(* IEC 61131-3 sources: JingjiangArm/moonboxpro_arm_8.4/Application/Application/任务列表/CommTask/轴号站号处理, 8 files *)

(* ---- KS_CheckArcIdValid.st ---- *)
(*@CES
Name=KS_CheckArcIdValid
Type=FunctionBlock
TypeGuid=6f9dac99-8de1-4efc-8465-68ac443b7d08
Guid=246184da-21c6-48ff-adc4-5d24f4660108
HasDeclaration=True
HasImplementation=True
*)
{DECLARATION}
FUNCTION KS_CheckArcIdValid : BOOL
VAR_INPUT
	i_iAxisId:INT;(*轴id*)
	i_iArcId:INT;(*套色id@修改后的*)
	i_pabyColorIdCurrent: POINTER TO ARRAY [1..MAX_UNIT_NUM] OF BYTE;(*色组色序*)
END_VAR
VAR
	iN: INT;
	xValid:BOOL:=TRUE;(*默认是有效的*)
END_VAR

{IMPLEMENTATION}
IF i_pabyColorIdCurrent<>0 THEN
	IF i_iAxisId>1 AND i_iArcId>1 THEN
		FOR iN:=1 TO i_iAxisId-1 BY 1 DO(*检查修改的轴前面的轴套色id*)
			IF i_pabyColorIdCurrent^[iN]>1 THEN(**)
				IF i_iArcId>i_pabyColorIdCurrent^[iN] THEN(*新修改的比上面轴的大就行*);
				ELSE(*小于等于任何一个都认为是无效的*)
					xValid:=FALSE;
					EXIT;
				END_IF
			END_IF
		END_FOR
	END_IF
END_IF

KS_CheckArcIdValid:=xValid;

(* ---- KS_GetArcIdList.st ---- *)
(*@CES
Name=KS_GetArcIdList
Type=FunctionBlock
TypeGuid=6f9dac99-8de1-4efc-8465-68ac443b7d08
Guid=d22e29e8-5d32-4a53-8a83-de107a05006d
HasDeclaration=True
HasImplementation=True
*)
{DECLARATION}
FUNCTION KS_GetArcIdList : BOOL
VAR_INPUT
	i_xEn:BOOL;(*更新列表使能标志*)
	i_iGrpAxisNum_Pu: INT; (*系的轴数量*)
	i_aiGrpAxisList: ARRAY [1..MAX_UNIT_NUM] OF INT; (*系的轴列表|已经按照升序排列了*)
	i_paxArcEnSts_Bak:POINTER TO ARRAY [1..MAX_UNIT_NUM] OF BOOL;(*套色使能备份值|用于检查是否套色使能切换*)
	i_pabyArcId_Bak:POINTER TO ARRAY [1..MAX_UNIT_NUM] OF BYTE;(*备份套色id*)
	(*系套色轴个数@可以输入0*)
	i_piGrpArcAxisNum_Pu:POINTER TO INT;
	i_axLinkage: ARRAY [1..MAX_UNIT_NUM] OF BOOL;
	i_axThisUnitEna: ARRAY [1..MAX_UNIT_NUM] OF BOOL;
	i_axSwitchOn_CoatingPrn: ARRAY [1..MAX_UNIT_NUM] OF BOOL;
	i_pabyColorIdCurrent: POINTER TO ARRAY [1..MAX_UNIT_NUM] OF BYTE;(*色组色序*)

END_VAR
VAR
	iN:INT;
	iUnitId:INT;
	xArcEnSts:BOOL;(*套色使能值|用于检查是否套色使能切换*)
	axArcEnSts_Bak:ARRAY [1..MAX_UNIT_NUM] OF BOOL;(*套色使能备份值|用于检查是否套色使能切换*)
	abyArcId_Bak:ARRAY [1..MAX_UNIT_NUM] OF BYTE;(*备份套色id*)
	(*系套色个数*)
	iGrpArcAxisNum_Pu:INT;
	xNeedUpdate: BOOL;
	byAxisIdArcValid: BYTE;(*最后一个未更新套色id|有效的轴id*)
	iAxisIdSa_Update: INT;(*更新的起始id@后面轴的套色id都更新*)
	xArcIdLocked:BOOL;(*套色id被锁定了|在更新的时候不修改这个值*)
	xRtn: BOOL;
	xUpdateArcId_BakValue: BOOL;(*更新套色id的备份值*)
	iIndex: INT;
END_VAR

{IMPLEMENTATION}
IF i_paxArcEnSts_Bak<>0 AND
	i_pabyArcId_Bak<>0 AND
	i_pabyColorIdCurrent<>0 THEN

	IF i_xEn THEN
		axArcEnSts_Bak:=i_paxArcEnSts_Bak^;(*获取之前的备份值*)
		abyArcId_Bak:=i_pabyArcId_Bak^;(*备份套色id*)

		FOR iN:=1 TO i_iGrpAxisNum_Pu BY 1 DO
			iUnitId:=i_aiGrpAxisList[iN];

			xArcEnSts:=i_axThisUnitEna[iUnitId] AND(*使能了*)
				i_axLinkage[iUnitId] AND(*联动了*)
				(NOT i_axSwitchOn_CoatingPrn[iUnitId]);(*不是涂布色组*)

			IF xArcEnSts<>axArcEnSts_Bak[iUnitId] THEN(*有轴的状态发生变化了*)
				IF NOT xNeedUpdate THEN(*记录需要更新的开始轴id*)
					iAxisIdSa_Update:=iUnitId;
				END_IF
				xNeedUpdate:=TRUE;
			END_IF

			(*记录最后一个不更新套色id的轴*)
			IF NOT xNeedUpdate THEN(*还没找到需要变化的轴id*)
				IF i_pabyColorIdCurrent^[iUnitId]<>0 THEN
					byAxisIdArcValid:= i_pabyColorIdCurrent^[iUnitId];
				END_IF
			END_IF
			axArcEnSts_Bak[iUnitId]:=xArcEnSts;
		END_FOR

		IF NOT xNeedUpdate THEN(*手动更新列表@注意调用顺序*)
			FOR iN:=1 TO i_iGrpAxisNum_Pu BY 1 DO
				iUnitId:=i_aiGrpAxisList[iN];
				xArcEnSts:=axArcEnSts_Bak[iUnitId];
				IF NOT xArcEnSts THEN(*套色不使能的时候 手动也不能输入*)
					i_pabyColorIdCurrent^[iUnitId]:=0;(*强制写0*)
				ELSE
					IF i_pabyColorIdCurrent^[iUnitId]=0 THEN(*输入了0则强制写成备份值*)
						i_pabyColorIdCurrent^[iUnitId]:=abyArcId_Bak[iUnitId];
						EXIT;(*手动修改了*)
					ELSE
						IF abyArcId_Bak[iUnitId]<>i_pabyColorIdCurrent^[iUnitId] THEN(*id被修改了*)
							xRtn:=KS_CheckArcIdValid(iUnitId,i_pabyColorIdCurrent^[iUnitId],i_pabyColorIdCurrent);
							IF xRtn THEN(*id合法@手动修改成功了|后面的列表需要同步更新*)
								xNeedUpdate:=TRUE;(*由下面逻辑生成*)
								iAxisIdSa_Update:=iUnitId;
								byAxisIdArcValid:=i_pabyColorIdCurrent^[iUnitId]-1;(*更新的时候会+1*)
							ELSE(*不合法@保持之前的*)
								i_pabyColorIdCurrent^[iUnitId]:=abyArcId_Bak[iUnitId];
							END_IF
							(*pstStAxisParam^.byColorIdCurrent 界面修改的,不在同一个任务中,防止不能抓住改变的状态
							置标志只有进入过这里才更新备份值*)
							xUpdateArcId_BakValue:=TRUE;

							EXIT;(*手动修改了*)
						END_IF
					END_IF
				END_IF
			END_FOR
		END_IF

		(*上面执行完成后axArcEnSts_Bak 中存储的每个色组是否套色的状态*)
		IF xNeedUpdate THEN(*自动更新列表了*)
			(*套色轴个数初始化*)
			IF byAxisIdArcValid<>0 THEN
				iGrpArcAxisNum_Pu:=BYTE_TO_INT(byAxisIdArcValid);
			ELSE
				iGrpArcAxisNum_Pu:=0;
			END_IF

			(*找到起始轴的索引值*)
			FOR iN:=1 TO i_iGrpAxisNum_Pu BY 1 DO
				iUnitId:=i_aiGrpAxisList[iN];
				IF iAxisIdSa_Update = iUnitId THEN
					iIndex:=iN;
					EXIT;
				END_IF
			END_FOR

			FOR iN:=iIndex TO i_iGrpAxisNum_Pu BY 1 DO(*从变化的轴这里开始，更新后面的套色id*)
				iUnitId:=i_aiGrpAxisList[iN];
				xArcEnSts:=axArcEnSts_Bak[iUnitId];

//xArcIdLocked;(*还未处理*)

				IF xArcEnSts THEN(*套色使能了*)
					iGrpArcAxisNum_Pu:=iGrpArcAxisNum_Pu+1;
					IF NOT xArcIdLocked THEN(*套色Id未被锁定*)
						i_pabyColorIdCurrent^[iUnitId]:=INT_TO_BYTE(iGrpArcAxisNum_Pu);
					ELSE(*套色Id被锁定了|当前色序id不做修改,更新套色轴个数变量*)
						IF i_pabyColorIdCurrent^[iUnitId]>iGrpArcAxisNum_Pu THEN
							iGrpArcAxisNum_Pu:=i_pabyColorIdCurrent^[iUnitId];
						ELSE
							i_pabyColorIdCurrent^[iUnitId]:=INT_TO_BYTE(iGrpArcAxisNum_Pu);
						END_IF
					END_IF
				ELSE
					i_pabyColorIdCurrent^[iUnitId]:=0;
				END_IF
			END_FOR
		ELSE(*在不更新的时候支持手动的输入*);
		END_IF

		(*更新存储的备份值@不用做专门的备份值初始化,因为刚上电的大概率肯定会更新列表*)
		FOR iN:=1 TO i_iGrpAxisNum_Pu BY 1 DO
			iUnitId:=i_aiGrpAxisList[iN];
			(*pstStAxisParam^.byColorIdCurrent 界面修改的,不在同一个任务中,防止不能抓住改变的状态
			置标志只有进入过上面逻辑更新备份值*)
			IF xUpdateArcId_BakValue OR xNeedUpdate THEN(*或者更新了列表后就更新*)
				abyArcId_Bak[iUnitId]:=i_pabyColorIdCurrent^[iUnitId];
			END_IF
		END_FOR
	ELSE;(*不使能*)
	END_IF

	i_paxArcEnSts_Bak^:=axArcEnSts_Bak;(*更新备份值|en=false 全部写成false*)
	i_pabyArcId_Bak^:=abyArcId_Bak;(*备份套色id*)
END_IF

IF i_piGrpArcAxisNum_Pu<>0 THEN
	i_piGrpArcAxisNum_Pu^:=iGrpArcAxisNum_Pu;
END_IF

(* ---- KS_GetAxisIdByStationId.st ---- *)
(*@CES
Name=KS_GetAxisIdByStationId
Type=FunctionBlock
TypeGuid=6f9dac99-8de1-4efc-8465-68ac443b7d08
Guid=70bbd18d-dc05-4e5d-8cd8-b579d4b6dda1
HasDeclaration=True
HasImplementation=True
*)
{DECLARATION}
FUNCTION KS_GetAxisIdByStationId : INT
VAR_INPUT
 	i_StationId: INT;
	i_aiStationList_UnitController: ARRAY [1..MAX_STATION_NUM] OF INT;(*用月光宝盒/PRO时候，需要一个控制器列表，用于通讯？*)
END_VAR
VAR
	iUnitId:INT;
	iN:INT;
	xResult: BOOL;
END_VAR

{IMPLEMENTATION}
iUnitId := 0;
IF i_StationId>=0 AND i_StationId<= MAX_STATION_NUM THEN
	FOR iN := 1 TO MAX_STATION_NUM BY 1 DO
		IF i_aiStationList_UnitController[iN] = i_StationId THEN
			iUnitId := iN;
			EXIT;
		END_IF
	END_FOR
END_IF
KS_GetAxisIdByStationId := iUnitId;

(* ---- KS_GetCoreAndAxisIdByStationId.st ---- *)
(*@CES
Name=KS_GetCoreAndAxisIdByStationId
Type=FunctionBlock
TypeGuid=6f9dac99-8de1-4efc-8465-68ac443b7d08
Guid=a5371cf2-ec50-4947-b43a-b8c7da498013
HasDeclaration=True
HasImplementation=True
*)
{DECLARATION}
FUNCTION KS_GetCoreAndAxisIdByStationId : INT
VAR_INPUT
	i_StationId: INT;
	i_piCoreId: POINTER TO INT;
	i_piAxisId: POINTER TO INT;
	i_aiStationIdList						: ARRAY [1..MAX_STATION_NUM] OF INT;(* 站号列表 *)
END_VAR
VAR
	iCoreId:INT;
	iUnitId:INT;
	iN:INT;
	xResult: BOOL;
END_VAR

{IMPLEMENTATION}
xResult := 0;
IF i_StationId>=0 AND i_StationId<= MAX_STATION_NUM AND
	i_piCoreId <>0 AND i_piAxisId <> 0 THEN

	FOR iN := 1 TO MAX_STATION_NUM BY 1 DO
		IF i_aiStationIdList[iN] = i_StationId THEN
			iUnitId := iN;
			EXIT;
		END_IF
	END_FOR
	IF iUnitId > 64 THEN
		iCoreId := 2;
		iUnitId := iUnitId - 64;
	ELSE
		iCoreId := 1;
	END_IF
	i_piCoreId^ := iCoreId;
	i_piAxisId^ := iUnitId;
END_IF

(* ---- KS_GetGrpIdByAxisId.st ---- *)
(*@CES
Name=KS_GetGrpIdByAxisId
Type=FunctionBlock
TypeGuid=6f9dac99-8de1-4efc-8465-68ac443b7d08
Guid=12f92d96-019f-4162-be83-866401d8db4e
HasDeclaration=True
HasImplementation=True
*)
{DECLARATION}
FUNCTION KS_GetGrpIdByAxisId : INT(*-1:参数错误或无效; 1=A系; 2=B系;|*)
VAR_INPUT
	i_iAxisId: INT; (* 轴id *)
	i_pstStSysParam: POINTER TO StSysParam; (* 参数 *)
	i_piAxisTypeId: POINTER TO INT := 0; (* 轴类型/0色组/1放牵/2收牵/3放料/4收料 *)
END_VAR
VAR
	iResult: INT;
	iUMax: INT;
	xDualUwRw: BOOL;
	xAsOneMachine: BOOL;
	pstStUnitParam_Save: POINTER TO StUnitParam_Save;
	xUwRwByServo: BOOL; (* 2021.1.14.222029/收放料采用伺服控制 *)
END_VAR
{IMPLEMENTATION}
iResult:= -1;
IF i_piAxisTypeId<>0 THEN
	i_piAxisTypeId^:= 0;
END_IF
IF (i_iAxisId>=1 AND i_iAxisId<=MAX_STATION_NUM) AND
	i_pstStSysParam<>0 THEN
	(*the parameters are valid|*)

	pstStUnitParam_Save:= ADR(i_pstStSysParam^.astStUnitParam_Save[i_iAxisId]);(*轴入口地址|*)

	iUMax:= i_pstStSysParam^.stStSysParam_Save.iUnitMaxNum;(*最大机组数|*)
	xDualUwRw:= i_pstStSysParam^.stStSysParam_Save.dwEquipmentProf.20;(*双收双放|*)
	xAsOneMachine:= i_pstStSysParam^.stStSysParam_Save.dwEquipmentProf.21;(*A放B收|*)
	xUwRwByServo:= i_pstStSysParam^.stStSysParam_Save.dwEquipmentProf.22; (* 2021.1.14.222103|收放料伺服控制 *)

	IF i_iAxisId>iUMax THEN
		(*牵引*)
		(*或者收放料|2021.1.14.222215 *)
		IF xDualUwRw THEN(*双收双放|*)
			IF xAsOneMachine THEN(*当整台开|*)
				CASE i_iAxisId OF
				31,32:
					iResult:= 1;(*只有A系|*)
					IF i_piAxisTypeId<>0 AND i_iAxisId=31 THEN
						i_piAxisTypeId^:= 1;(*放牵|*)
					ELSIF i_piAxisTypeId<>0 AND i_iAxisId=32 THEN
						i_piAxisTypeId^:= 2;(*收牵|*)
					END_IF
				25,26,27,28: (* 2021.1.14.223803/扩展的类型 *)
					IF xUwRwByServo THEN
						iResult:= 1; (* 只有A系 *)
						IF i_piAxisTypeId<>0 AND (i_iAxisId=25 OR i_iAxisId=26) THEN (* 放料 *)
							i_piAxisTypeId^:= 3; (* 放料 *)
						ELSIF i_piAxisTypeId<>0 AND (i_iAxisId=27 OR i_iAxisId=28) THEN (* 收料 *)
							i_piAxisTypeId^:= 4; (* 收料 *)
						END_IF
					END_IF
				ELSE;
				END_CASE
			ELSE
				(*分A/B系*)
				CASE i_iAxisId OF
				30,31:
					iResult:= 1;(*A系|*)
					IF i_piAxisTypeId<>0 AND i_iAxisId=31 THEN
						i_piAxisTypeId^:= 1;(*放牵|*)
					ELSIF i_piAxisTypeId<>0 AND i_iAxisId=30 THEN
						i_piAxisTypeId^:= 2;(*收牵|*)
					END_IF
				29,32:
					iResult:= 2;(*B系|*)
					IF i_piAxisTypeId<>0 AND i_iAxisId=29 THEN
						i_piAxisTypeId^:= 1;(*放牵|*)
					ELSIF i_piAxisTypeId<>0 AND i_iAxisId=32 THEN
						i_piAxisTypeId^:= 2;(*收牵|*)
					END_IF
				23,24,25,26: (* 2021.1.14.222755/扩展 *)
					IF xUwRwByServo THEN
						iResult:= 1; (* A系 *)
						IF i_piAxisTypeId<>0 AND (i_iAxisId=25 OR i_iAxisId=26) THEN (* 放料 *)
							i_piAxisTypeId^:= 3; (* 放料 *)
						ELSIF i_piAxisTypeId<>0 AND (i_iAxisId=23 OR i_iAxisId=24) THEN (* 收料 *)
							i_piAxisTypeId^:= 4; (* 收料 *)
						END_IF
					END_IF
				21,22,27,28: (* 2021.1.14.222755/扩展 *)
					IF xUwRwByServo THEN
						iResult:= 2; (* B系 *)
						IF i_piAxisTypeId<>0 AND (i_iAxisId=21 OR i_iAxisId=22) THEN (* 放料 *)
							i_piAxisTypeId^:= 3; (* 放料 *)
						ELSIF i_piAxisTypeId<>0 AND (i_iAxisId=27 OR i_iAxisId=28) THEN (* 收料 *)
							i_piAxisTypeId^:= 4; (* 收料 *)
						END_IF
					END_IF
				ELSE;
				END_CASE
			END_IF
		ELSE(*标准机型*)
			iResult:= 1;(*只有A系|*)
			IF i_piAxisTypeId<>0 AND i_iAxisId=31 THEN
				i_piAxisTypeId^:= 1;(*放牵|*)
			ELSIF i_piAxisTypeId<>0 AND i_iAxisId=32 THEN
				i_piAxisTypeId^:= 2;(*收牵|*)
			ELSIF i_piAxisTypeId<>0 AND xUwRwByServo AND (i_iAxisId=25 OR i_iAxisId=26) THEN (* 2021.1.14.222755/放料 *)
				i_piAxisTypeId^:= 3; (* 放料 *)
			ELSIF i_piAxisTypeId<>0 AND xUwRwByServo AND (i_iAxisId=27 OR i_iAxisId=28) THEN (* 2021.1.14.222755/收料 *)
				i_piAxisTypeId^:= 4; (* 收料 *)
			END_IF
		END_IF
	ELSE
		(*色组*)
		IF xDualUwRw AND (NOT xAsOneMachine) THEN(*双收双放且不作为单台印刷机开*)
			IF pstStUnitParam_Save^.byGrpId=1 OR pstStUnitParam_Save^.byGrpId=2 THEN
				;
			ELSE(*如果系id有问题就都分配到A系|*)
				pstStUnitParam_Save^.byGrpId:= 1;
			END_IF
		ELSE
			pstStUnitParam_Save^.byGrpId:= 1;
		END_IF
		iResult:= BYTE_TO_INT(pstStUnitParam_Save^.byGrpId);
	END_IF
END_IF

KS_GetGrpIdByAxisId:= iResult;

(* ---- KS_GetUnitIdAndTypeByStationId.st ---- *)
(*@CES
Name=KS_GetUnitIdAndTypeByStationId
Type=FunctionBlock
TypeGuid=6f9dac99-8de1-4efc-8465-68ac443b7d08
Guid=562049e6-f238-457e-b203-3358a7713818
HasDeclaration=True
HasImplementation=True
*)
{DECLARATION}
FUNCTION KS_GetUnitIdAndTypeByStationId : bool
VAR_INPUT
	i_StationId: INT;
	i_piUnitId: POINTER TO INT;
	i_piTypeId: POINTER TO INT;
	i_pstStSysCfgStruct: POINTER TO StSysCfgStruct;
END_VAR
VAR
	iUnitId:INT;
	iTypeId:INT;
	iN:INT;
	xResult: BOOL;
END_VAR

{IMPLEMENTATION}
(*	OBJ_IS_UNDEFINED,
	OBJ_IS_UNWIND_A,(* 放卷A *)
	OBJ_IS_UNWIND_B,(* 放卷B *)
	OBJ_IS_REWIND_A,(* 收卷A *)
	OBJ_IS_REWIND_B,(* 收卷B *)
	OBJ_IS_INFEED,(* 放牵 *)
	OBJ_IS_OUTFEED,(* 收牵 *)
	OBJ_IS_BOTTOM_ROLLER,(* 色组底辊 *)
	OBJ_IS_PRN_ROLLER,(* 色组版辊 *)
	OBJ_IS_NET_ROLLER,(* 色组网辊 *)
	OBJ_IS_PRN_ROLLER_PRESSURE_M,(* 色组版辊压力M侧 *)
////OBJ_IS_PRN_ROLLER_PRESSURE_G,(* 色组版辊压力G侧 *)
////OBJ_IS_NET_ROLLER_PRESSURE_M,(* 色组网辊压力M侧 *)
////OBJ_IS_NET_ROLLER_PRESSURE_G,(* 色组网辊压力G侧 *)
////OBJ_IS_HORIZ_MOTION,(* 横向运动电机/2022.6.8.142000 *)
////OBJ_IS_CENTRAL_DRUM(* 中心滚筒/2022.6.8.135513 *)*)
xResult:= FALSE;
IF i_StationId>=0 AND i_StationId<= MAX_STATION_NUM AND
	i_pstStSysCfgStruct<>0 THEN
	IF i_pstStSysCfgStruct^.stStAxisCfgStruct_IF_I.iSid=i_StationId AND i_pstStSysCfgStruct^.stStAxisCfgStruct_IF_I.dwAxisProf.0 THEN
		iUnitId:= 31;
		iTypeId:= OBJ_IS_INFEED;
	ELSIF i_pstStSysCfgStruct^.stStAxisCfgStruct_OF_I.iSid=i_StationId AND i_pstStSysCfgStruct^.stStAxisCfgStruct_OF_I.dwAxisProf.0 THEN
		iUnitId:= 32;
		iTypeId:= OBJ_IS_OUTFEED;
	ELSIF i_pstStSysCfgStruct^.astStAxisCfgStruct_UW_I[1].iSid=i_StationId AND i_pstStSysCfgStruct^.astStAxisCfgStruct_UW_I[1].dwAxisProf.0 THEN
		iUnitId:= 25;
		iTypeId:= OBJ_IS_UNWIND_A;
	ELSIF i_pstStSysCfgStruct^.astStAxisCfgStruct_UW_I[2].iSid=i_StationId AND i_pstStSysCfgStruct^.astStAxisCfgStruct_UW_I[2].dwAxisProf.0 THEN
		iUnitId:= 26;
		iTypeId:= OBJ_IS_UNWIND_B;
	ELSIF i_pstStSysCfgStruct^.astStAxisCfgStruct_RW_I[1].iSid=i_StationId AND i_pstStSysCfgStruct^.astStAxisCfgStruct_RW_I[1].dwAxisProf.0 THEN
		iUnitId:= 27;
		iTypeId:= OBJ_IS_REWIND_A;
	ELSIF i_pstStSysCfgStruct^.astStAxisCfgStruct_RW_I[2].iSid=i_StationId AND i_pstStSysCfgStruct^.astStAxisCfgStruct_RW_I[2].dwAxisProf.0 THEN
		iUnitId:= 28;
		iTypeId:= OBJ_IS_REWIND_B;
	ELSIF i_pstStSysCfgStruct^.astStAxisCfgStruct_CD_i[1].iSid=i_StationId AND i_pstStSysCfgStruct^.astStAxisCfgStruct_CD_I[1].dwAxisProf.0 THEN
		iUnitId:= 20;(*中心辊增加一个|2024.04.01.094732*)
		iTypeId:= OBJ_IS_CENTRAL_DRUM;
	ELSIF i_pstStSysCfgStruct^.astStAxisCfgStruct_CD_i[2].iSid=i_StationId AND i_pstStSysCfgStruct^.astStAxisCfgStruct_CD_I[2].dwAxisProf.0 THEN
		iUnitId:= 21;(*中心辊增加一个|2024.04.01.094732*)
		iTypeId:= OBJ_IS_CENTRAL_DRUM;
	ELSE
		FOR iN:=1 TO MAX_UNIT_NUM BY 1 DO
			IF i_pstStSysCfgStruct^.astStAxisCfgStruct_PR_[iN].iSid= i_StationId AND i_pstStSysCfgStruct^.astStAxisCfgStruct_PR_[iN].dwAxisProf.0 THEN
				iUnitId:= iN;
				iTypeId:= OBJ_IS_PRN_ROLLER;
			ELSIF i_pstStSysCfgStruct^.astStAxisCfgStruct_NR_[iN].iSid= i_StationId AND i_pstStSysCfgStruct^.astStAxisCfgStruct_NR_[iN].dwAxisProf.0 THEN
				iUnitId:= iN;
				iTypeId:= OBJ_IS_NET_ROLLER;
			ELSIF i_pstStSysCfgStruct^.astStAxisCfgStruct_BR_[iN].iSid= i_StationId AND i_pstStSysCfgStruct^.astStAxisCfgStruct_BR_[iN].dwAxisProf.0 THEN
				iUnitId:= iN;
				iTypeId:= OBJ_IS_BOTTOM_ROLLER;
			ELSIF i_pstStSysCfgStruct^.astStAxisCfgStruct_HORIZ_[iN].iSid= i_StationId AND i_pstStSysCfgStruct^.astStAxisCfgStruct_HORIZ_[iN].dwAxisProf.0 THEN
				iUnitId:= iN;
				iTypeId:= OBJ_IS_HORIZ_MOTION;
			ELSIF i_pstStSysCfgStruct^.astStAxisCfgStruct_PR_M_[iN].iSid= i_StationId AND i_pstStSysCfgStruct^.astStAxisCfgStruct_PR_M_[iN].dwAxisProf.0 THEN
				iUnitId:= iN;
				iTypeId:= OBJ_IS_PRN_ROLLER_PRESSURE_M;
			ELSIF i_pstStSysCfgStruct^.astStAxisCfgStruct_PR_G_[iN].iSid= i_StationId AND i_pstStSysCfgStruct^.astStAxisCfgStruct_PR_G_[iN].dwAxisProf.0 THEN
				iUnitId:= iN;
				iTypeId:= OBJ_IS_PRN_ROLLER_PRESSURE_G;
			ELSIF i_pstStSysCfgStruct^.astStAxisCfgStruct_NR_M_[iN].iSid= i_StationId AND i_pstStSysCfgStruct^.astStAxisCfgStruct_NR_M_[iN].dwAxisProf.0 THEN
				iUnitId:= iN;
				iTypeId:= OBJ_IS_NET_ROLLER_PRESSURE_M;
			ELSIF i_pstStSysCfgStruct^.astStAxisCfgStruct_NR_G_[iN].iSid= i_StationId AND i_pstStSysCfgStruct^.astStAxisCfgStruct_NR_G_[iN].dwAxisProf.0 THEN
				iUnitId:= iN;
				iTypeId:= OBJ_IS_NET_ROLLER_PRESSURE_G;
			ELSIF i_pstStSysCfgStruct^.astStAxisCfgStruct_PC_[iN].iSid=i_StationId AND i_pstStSysCfgStruct^.astStAxisCfgStruct_PC_[iN].dwAxisProf.0 THEN
				iUnitId:= iN;(*光电眼行走机构 | 2024.04.01.092649*)
				iTypeId:= OBJ_IS_PHOTOCELL;
			ELSIF i_pstStSysCfgStruct^.astStAxisCfgStruct_STR_M_[iN].iSid= i_StationId AND i_pstStSysCfgStruct^.astStAxisCfgStruct_STR_M_[iN].dwAxisProf.0 THEN
				iUnitId:= iN;
				iTypeId:= OBJ_IS_STR_ROLLER_PRESSURE_M;
			ELSIF i_pstStSysCfgStruct^.astStAxisCfgStruct_STR_G_[iN].iSid= i_StationId AND i_pstStSysCfgStruct^.astStAxisCfgStruct_STR_G_[iN].dwAxisProf.0 THEN
				iUnitId:= iN;
				iTypeId:= OBJ_IS_STR_ROLLER_PRESSURE_G;
			END_IF
		END_FOR
	END_IF

	IF i_piUnitId<>0 THEN
		i_piUnitId^:= iUnitId;
	END_IF
	IF i_piTypeId<>0 THEN
		i_piTypeId^:= iTypeId;
	END_IF
END_IF

KS_GetUnitIdAndTypeByStationId:= xResult;

(* ---- KS_IsValidStationNR.st ---- *)
(*@CES
Name=KS_IsValidStationNR
Type=FunctionBlock
TypeGuid=6f9dac99-8de1-4efc-8465-68ac443b7d08
Guid=c4580633-d047-4a45-9578-afb5bd290b41
HasDeclaration=True
HasImplementation=True
*)
{DECLARATION}
FUNCTION KS_IsValidStationNR : BOOL
VAR_INPUT
	i_iStationNR: INT;
END_VAR
VAR
	xResult: BOOL;
END_VAR

{IMPLEMENTATION}
IF i_iStationNR>=0 AND i_iStationNR<MAX_STATION_NUM THEN
	xResult:= TRUE;
ELSE
	xResult:= FALSE;
END_IF
KS_IsValidStationNR:= xResult;

(* ---- KS_IsValidUnitNR.st ---- *)
(*@CES
Name=KS_IsValidUnitNR
Type=FunctionBlock
TypeGuid=6f9dac99-8de1-4efc-8465-68ac443b7d08
Guid=8ab37e44-6a25-425d-9d9c-1a5dcec00b7a
HasDeclaration=True
HasImplementation=True
*)
{DECLARATION}
FUNCTION KS_IsValidUnitNR : BOOL
VAR_INPUT
	i_iUnitNR: INT;
END_VAR
VAR
	xResult: BOOL;
END_VAR
{IMPLEMENTATION}
IF i_iUnitNR>=1 AND i_iUnitNR<=MAX_UNIT_NUM THEN
	xResult:= TRUE;
ELSE
	xResult:= FALSE;
END_IF
KS_IsValidUnitNR:= xResult;
